(* PLC project zarechnaya.project, CODESYS CODESYS V3.5 SP17 Patch 3 *)
(* stored: creationDateTime 2026-10-20T05:42:22.3967198, modificationDateTime 1601-01-01T03:00:00 *)

TYPE U_Status : UNION
  w : WORD;
  b : ARRAY[0..1] OF BYTE;
END_UNION;
END_TYPE
